Yaskawa INFORM job: HOME_MO.JBI

/JOB
//NAME HOME_MO
//POS
///NPOS 1,0,0,0,0,0
///TOOL 9
///POSTYPE PULSE
///PULSE
C00000=35,-55,-66,-180,-91,180
//INST
///DATE 2026/10/26 01:19
///COMM Generated using RoboDK
///ATTR SC,RW
///GROUP1 RB1
NOP
'Program generated by Vertical
'Bot Studio for Motoman ES200D
' on 25/10/2026 12:00:00
'Using nominal kinematics.
'Using Frame 1 (targets wrt ba
'se):
'1724.5,-1789.7,1123.6,0.0,0.0
',93.8
'Tool Spindle should be close
'to:
'417.9,0.0,132.0,0.0,90.0,0.0
MOVJ C00000 VJ=50.00
END
